(* IEC 61131-3 sources: codesys-to-s7/tests/corpus/C2S7-TYPE-ALIAS/pos, 1 file *)

(* ---- input.st ---- *)
TYPE T_Pct : INT; END_TYPE
FUNCTION_BLOCK FB_Case
VAR
    p : T_Pct;
END_VAR
p := 5;
END_FUNCTION_BLOCK
